Fanuc KAREL source: ka00109.KL

-- PROVISIONAL review KL for V770-1; original PC SHA256 b9177ca7e9fef1ba4756e717ed3ec298cdfa6a45fa42598ec440476d82e84ab0
-- Incomplete behavior may be omitted. Consult companion uncertainty JSON. Do not deploy.
PROGRAM KA00109
%NOLOCKGROUP
VAR
  DST : INTEGER
-- UNRESOLVED_DECL SRC type=00001c
BEGIN
  -- UNRESOLVED_PC offsets 5-15; opcodes 9D,22,A5
  -- UNRESOLVED_PC offsets 20-32; opcodes 21,23
  -- UNRESOLVED_PC offsets 37-41; opcodes 7F
END KA00109
